SUBAPPLICATION doppeltwirkend (* Subapplication Type *)
  (* Standard: 61499-2 *)
  (* Version 1.0, 2023-01-29, Franz *)
  IMPORT logiBUS::io::DQ::logiBUS_DO::Invalid;
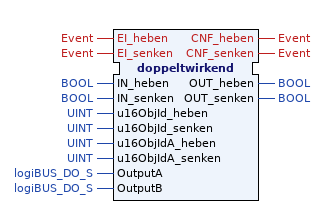
  EVENT_INPUT
    EI_heben;
    EI_senken;
  END_EVENT
  EVENT_OUTPUT
    CNF_heben;
    CNF_senken;
  END_EVENT
  VAR_INPUT
    IN_heben : BOOL;
    IN_senken : BOOL;
    u16ObjId_heben : UINT;
    u16ObjId_senken : UINT;
    u16ObjIdA_heben : UINT;
    u16ObjIdA_senken : UINT;
    OutputA : logiBUS::io::DQ::logiBUS_DO_S := Invalid;
    OutputB : logiBUS::io::DQ::logiBUS_DO_S := Invalid;
  END_VAR
  VAR_OUTPUT
    OUT_heben : BOOL;
    OUT_senken : BOOL;
  END_VAR
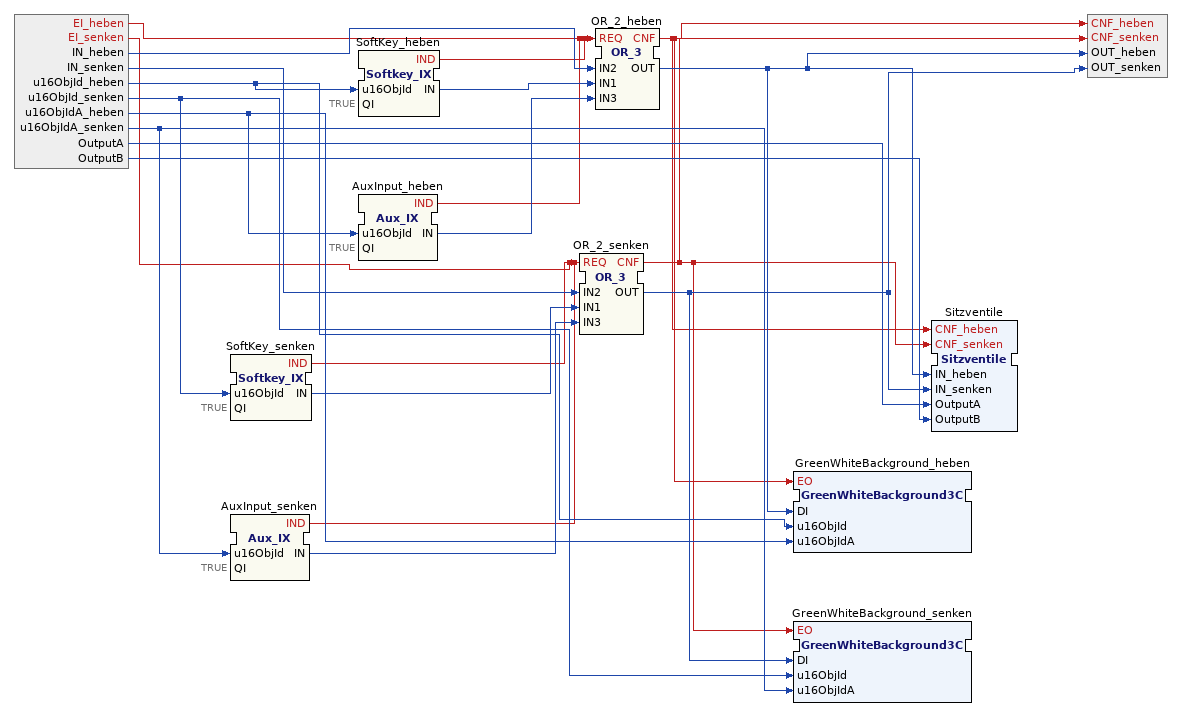
  FBS
    OR_2_heben : iec61131::bitwiseOperators::OR_3;
    OR_2_senken : iec61131::bitwiseOperators::OR_3;
    SoftKey_heben : isobus::UT::io::Softkey::Softkey_IX(QI := TRUE);
    AuxInput_heben : isobus::UT::io::Auxiliary::IN::Aux_IX(QI := TRUE);
    SoftKey_senken : isobus::UT::io::Softkey::Softkey_IX(QI := TRUE);
    AuxInput_senken : isobus::UT::io::Auxiliary::IN::Aux_IX(QI := TRUE);
  END_FBS
  SUBAPPS
    GreenWhiteBackground_heben : MyLib::sys::GreenWhiteBackground3C;
    GreenWhiteBackground_senken : MyLib::sys::GreenWhiteBackground3C;
    Sitzventile : Sitzventile;
  END_SUBAPPS
  EVENT_CONNECTIONS
    EI_heben TO OR_2_heben.REQ;
    OR_2_heben.CNF TO CNF_heben;
    EI_senken TO OR_2_senken.REQ;
    OR_2_senken.CNF TO CNF_senken;
    OR_2_heben.CNF TO GreenWhiteBackground_heben.EO;
    OR_2_senken.CNF TO GreenWhiteBackground_senken.EO;
    OR_2_heben.CNF TO Sitzventile.CNF_heben;
    OR_2_senken.CNF TO Sitzventile.CNF_senken;
    SoftKey_heben.IND TO OR_2_heben.REQ;
    AuxInput_heben.IND TO OR_2_heben.REQ;
    SoftKey_senken.IND TO OR_2_senken.REQ;
    AuxInput_senken.IND TO OR_2_senken.REQ;
  END_CONNECTIONS
  DATA_CONNECTIONS
    OutputB TO Sitzventile.OutputB;
    OutputA TO Sitzventile.OutputA;
    u16ObjIdA_senken TO AuxInput_senken.u16ObjId;
    u16ObjIdA_heben TO AuxInput_heben.u16ObjId;
    u16ObjId_heben TO SoftKey_heben.u16ObjId;
    u16ObjId_senken TO SoftKey_senken.u16ObjId;
    IN_heben TO OR_2_heben.IN2;
    OR_2_heben.OUT TO OUT_heben;
    IN_senken TO OR_2_senken.IN2;
    OR_2_senken.OUT TO OUT_senken;
    OR_2_heben.OUT TO GreenWhiteBackground_heben.DI;
    OR_2_senken.OUT TO GreenWhiteBackground_senken.DI;
    u16ObjId_heben TO GreenWhiteBackground_heben.u16ObjId;
    u16ObjId_senken TO GreenWhiteBackground_senken.u16ObjId;
    u16ObjIdA_heben TO GreenWhiteBackground_heben.u16ObjIdA;
    u16ObjIdA_senken TO GreenWhiteBackground_senken.u16ObjIdA;
    OR_2_heben.OUT TO Sitzventile.IN_heben;
    OR_2_senken.OUT TO Sitzventile.IN_senken;
    SoftKey_heben.IN TO OR_2_heben.IN1;
    AuxInput_heben.IN TO OR_2_heben.IN3;
    SoftKey_senken.IN TO OR_2_senken.IN1;
    AuxInput_senken.IN TO OR_2_senken.IN3;
  END_CONNECTIONS
END_SUBAPPLICATION
